// TIA Portal V21 export
// export: Created 2026-11-08T21:43:42.1133172Z, ExportSetting WithDefaults, DisplayName Totally Integrated Automation Portal, DisplayVersion V21 Update 3, DisplayName STEP 7 Professional, DisplayVersion V21 Update 3, DisplayName STEP 7 Safety, DisplayVersion V21, DisplayName Tech WebApplication, DisplayVersion V21, DisplayName WinCC Basic/Comfort/Advanced, DisplayVersion V21 Update 3, DisplayName WinCC Unified, DisplayVersion V21 Update 3
FUNCTION_BLOCK "FB_GraphEvt"   // FB77, GRAPH
VERSION : 0.1
// stored: AcknowledgeErrorsRequired true, AutoNumber true, GraphVersion 6.0, InitialValuesAcquisition false, IsIECCheckEnabled false, LanguageInNetworks LAD, LockOperatingMode false, PermanentILProcessingInMANMode false, SetENOAutomatically false, SkipSteps false, UDAEnableTagReadback false, WithAlarmHandling true
   // inherited from GRAPH_BASE
   VAR
      OFF_SQ_BASE : Bool;
   END_VAR
   VAR_INPUT
      OFF_SQ : Bool := false;   // Turn sequence off
      INIT_SQ : Bool := false;   // Set sequence to initial state
      ACK_EF : Bool := false;   // Acknowledge all errors and faults
      go : Bool;
      "a" : Bool;
      "b" : Bool;
      sv : Bool;
   END_VAR
   VAR_OUTPUT
      q1 : Bool;
      q2 : Bool;
      q3 : Bool;
   END_VAR
BEGIN
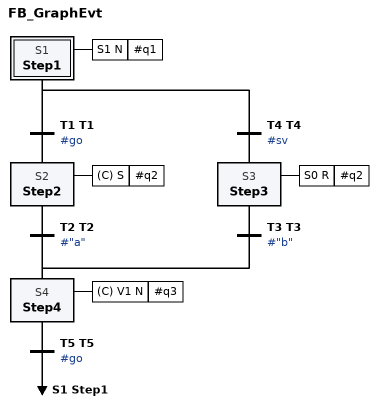
   // sequencer 1
   INITIAL_STEP Step1:   // S1, max time T#10S, warning time T#7S
      supervision V := #sv;
          S1  N    #q1
   END_STEP
   TRANSITION T1 FROM Step1 TO Step2   // T1
      := #go;
   END_TRANSITION
   TRANSITION T4 FROM Step1 TO Step3   // T4
      := #sv;
   END_TRANSITION
   STEP Step2:   // S2, max time T#10S, warning time T#7S
      supervision V := #sv;
      (C)     S    #q2
   END_STEP
   TRANSITION T2 FROM Step2 TO Step4   // T2
      := #"a";
   END_TRANSITION
   STEP Step3:   // S3, max time T#10S, warning time T#7S
      supervision V := #sv;
          S0  R    #q2
   END_STEP
   TRANSITION T3 FROM Step3 TO Step4   // T3
      := #"b";
   END_TRANSITION
   STEP Step4:   // S4, max time T#10S, warning time T#7S
      supervision V := #sv;
      (C) V1  N    #q3
   END_STEP
   TRANSITION T5 FROM Step4 TO Step1   // T5, jump
      := #go;
   END_TRANSITION
END_FUNCTION_BLOCK
